Staubli VAL3: copy.pgx

program copy()
  local string l_sMsg
  local string l_sInputName
  local bool l_bResult
  local bool l_bResult1
  local num l_nID
  local num l_i
  local bool l_bFound
  local num l_nSize
  local string l_sHeader
begin
  l_sMsg="复制"+sSelTraj+"到："
  l_bResult=userPagePrompt(l_sMsg,l_sInputName)
  if l_bResult
    call trajectory:isDefine(l_sInputName,l_bResult1)
    if !l_bResult1
      call trajectory:getSize(l_nSize)
      call getTrajID()
      l_nID=0
      do
        l_i=0
        do
          if l_nID==nIDIsExit[l_i]
            l_bFound=true
            l_nID=l_nID+1
          else
            l_bFound=false
          endIf
          l_i=l_i+1
        until l_bFound==false or l_i>=size(nIDIsExit)

      until l_bFound==false

      if l_nSize<10
        l_sHeader="0"+toString("",l_nID)+" "+l_sInputName
      else
        l_sHeader=toString("",l_nID)+" "+l_sInputName
      endIf

      call trajectory:copy(sSelTraj,l_sHeader,bToSave)
      call trajectory:onSave(bToSave)
    else
      userPageAlert("输入的名称重复！")
    endIf
  endIf
end
